TYPE ET_Gr01Home :
(
	ET_Gr01Home_eWaitExecute := 0,
	ET_Gr01Home_eWaitAxisStatus,
	ET_Gr01Home_eGetProcessPara,
	ET_Gr01Home_eSawbandStop,
	ET_Gr01Home_eWfSawbandStopped,
	ET_Gr01Home_eAxisSawbandGuide,
	ET_Gr01Home_eWfAxisSawbandGuide,
	ET_Gr01Home_eAxisSawBow,
	ET_Gr01Home_eWfAxisSawBow,
	ET_Gr01Home_eAxisAngle,
	ET_Gr01Home_eWfAxisAngle,
	ET_Gr01Home_eWfFreeToMove,
	ET_Gr01Home_eAxisSawBowMoveHomePos,
	ET_Gr01Home_eWfAxisSawBowInHomePos,
	ET_Gr01Home_eDone := 197,
	ET_Gr01Home_eError := 198,
	ET_Gr01Home_eNoExecute := 199
);
END_TYPE

(* stored: Version 1.1.0.1, ProductVersion 3.1.4024.15
   DUT ET_Gr01Home: Id {c7643085-5345-4161-9908-4c6f07a8f68d} *)
